// TIA Portal V19 export
DATA_BLOCK "SOLVENT_ADDITION_START"   // DB10
// stored: InstanceOfName START, InstanceOfType FB
"START"
   // VAR_INPUT
   //    RUNNING : Bool;
   // END_VAR
   // VAR_OUTPUT
   //    START_CMD : Bool;
   //    STOP_CMD : Bool;
   // END_VAR
   // VAR_IN_OUT
   //    "START/STOP" : Bool;
   // END_VAR
   // VAR
   //    START_PLS : Bool;
   //    IEC_Timer_0_Instance { S7_SetPoint := 'True'} : TOF_TIME;
   //    STOP_PLS : Bool;
   //    IEC_Timer_0_Instance_1 { S7_SetPoint := 'True'} : TOF_TIME;
   //    RUNNING_PLS : Bool;
   // END_VAR
BEGIN
END_DATA_BLOCK
